(* IEC 61131-3 sources: codesys-motor-control-station/src, 9 files *)

(* ---- types_and_globals.st ---- *)
// ===== E_FaultCode =====

{attribute 'qualified_only'}
{attribute 'strict'}
TYPE E_FaultCode :
(
    NONE     := 0,
    ESTOP    := 1,   // Emergency stop pressed or circuit broken
    OVERLOAD := 2    // Thermal overload relay tripped
) UINT;
END_TYPE

{attribute 'qualified_only'}
{attribute 'strict'}
TYPE E_FaultCode :
(
    NONE     := 0,
    ESTOP    := 1,   // Emergency stop pressed or circuit broken
    OVERLOAD := 2    // Thermal overload relay tripped
) UINT;
END_TYPE

// ===== E_StationState =====

{attribute 'qualified_only'}
{attribute 'strict'}
TYPE E_StationState :
(
    IDLE     := 0,   // Stopped, ready to start
    STARTING := 1,   // Soft-start ramp running
    RUNNING  := 2,   // At speed setpoint
    STOPPING := 3,   // Soft-stop ramp running
    FAULT    := 4    // Fault latched, outputs off
) UINT;
END_TYPE

// ===== ST_Config =====

TYPE ST_Config :
STRUCT
    tRampUp           : TIME := T#5S;    // Soft-start duration (0 Hz to setpoint)
    tRampDown         : TIME := T#5S;    // Soft-stop duration (setpoint to 0 Hz)
    rSpeedMin_Hz      : REAL := 5.0;     // Lowest allowed setpoint
    rSpeedMax_Hz      : REAL := 50.0;    // Highest allowed setpoint
    rSpeedSetpoint_Hz : REAL := 40.0;    // Operator target speed
END_STRUCT
END_TYPE

// ===== GVL_HMI =====

{attribute 'qualified_only'}
VAR_GLOBAL
    xStart        : BOOL;   // Momentary: TRUE while START is pressed
    xStop         : BOOL;   // Momentary: TRUE while STOP is pressed
    xReset        : BOOL;   // Momentary: TRUE while RESET is pressed
    xEStop        : BOOL;   // Latching switch: TRUE = E-stop pressed
    xOverloadTrip : BOOL;   // Latching switch: TRUE = overload tripped
    xSetpointUp   : BOOL;   // Momentary: setpoint +5 Hz
    xSetpointDown : BOOL;   // Momentary: setpoint -5 Hz
END_VAR

// ===== GVL_IO =====

{attribute 'qualified_only'}
VAR_GLOBAL
    // ---------- Inputs ----------
    iEStop_OK       : BOOL;   // NC contact: TRUE = healthy, FALSE = E-stop pressed or wire broken
    iStop_PB        : BOOL;   // NC contact: TRUE = released, FALSE = pressed
    iStart_PB       : BOOL;   // NO contact: TRUE = pressed
    iOverload_OK    : BOOL;   // NC contact: TRUE = healthy, FALSE = overload tripped
    iFaultReset_PB  : BOOL;   // NO contact: TRUE = pressed

    // ---------- Outputs ----------
    qContactor_KM1  : BOOL;   // Main contactor coil
    qDriveRun       : BOOL;   // Run command to the VFD
    qSpeedRef_Hz    : REAL;   // Speed reference sent to the VFD (analog output, in Hz)
    qLamp_Ready     : BOOL;   // White: station ready
    qLamp_Run       : BOOL;   // Green: motor running or ramping
    qLamp_Fault     : BOOL;   // Red: fault latched
END_VAR

// ===== GVL_SIM =====

{attribute 'qualified_only'}
VAR_GLOBAL
    xEnable       : BOOL := TRUE;   // TRUE = simulation writes the GVL_IO inputs

    // Simulated input conditions
    xEStop_OK     : BOOL := TRUE;   // TRUE = E-stop circuit healthy
    xStop_PB      : BOOL := TRUE;   // TRUE = Stop button released
    xStart_PB     : BOOL := FALSE;  // TRUE = Start button pressed
    xOverload_OK  : BOOL := TRUE;   // TRUE = overload circuit healthy
    xFaultReset_PB : BOOL := FALSE; // TRUE = reset button pressed
END_VAR

// ===== GVL_STATION =====

{attribute 'qualified_only'}
VAR_GLOBAL
    stConfig       : ST_Config;                                  // Tunable parameters
    eState         : E_StationState := E_StationState.IDLE;      // Current state machine state
    eFault         : E_FaultCode    := E_FaultCode.NONE;         // Active fault cause
    xFaultLatched  : BOOL;                                       // TRUE until reset
    xSafeToRun     : BOOL;                                       // TRUE only when no fault and all safety inputs healthy
    xRunLatched    : BOOL;                                       // Start/stop seal-in memory
    rSpeedRef_Hz   : REAL;                                       // Ramp output (feeds qSpeedRef_Hz)
    xAtSetpoint    : BOOL;                                       // Ramp has reached the setpoint
    xAtZero        : BOOL;                                       // Ramp has reached 0 Hz
    rRunHours      : REAL;                                       // Run time in hours (for display)
END_VAR

VAR_GLOBAL PERSISTENT RETAIN
    nRunSeconds    : UDINT;                                      // Drive-on time in seconds, survives power cycles
END_VAR

(* ---- FB_RampGenerator.st ---- *)
FUNCTION_BLOCK FB_RampGenerator
VAR_INPUT
    xEnable    : BOOL;              // TRUE = ramp up to target and hold, FALSE = ramp down to 0 Hz
    xForceZero : BOOL;              // TRUE = output jumps to 0 Hz immediately (fault)
    rTarget_Hz : REAL;              // Speed to ramp up to
    tRampUp    : TIME;              // Time to go from 0 Hz to target
    tRampDown  : TIME;              // Time to go from target to 0 Hz
    tCycle     : TIME := T#10MS;    // Task cycle time (must match MainTask)
END_VAR
VAR_OUTPUT
    rOutput_Hz  : REAL;             // Ramped speed reference
    xAtSetpoint : BOOL;             // Enabled and output equals target
    xAtZero     : BOOL;             // Output is 0 Hz
END_VAR
VAR
    rTargetSafe : REAL;             // Target limited to 0 Hz or more
    rGoal       : REAL;             // Where the output is heading right now
    rStepUp     : REAL;             // Hz added per scan while accelerating
    rStepDown   : REAL;             // Hz removed per scan while decelerating
END_VAR
VAR CONSTANT
    rTolerance  : REAL := 0.001;    // Comparison tolerance in Hz
    rMinStep    : REAL := 0.001;    // Smallest allowed step, so a ramp always finishes
END_VAR

// ---------- 1. Goal ----------
rTargetSafe := MAX(rTarget_Hz, 0.0);

IF xEnable THEN
    rGoal := rTargetSafe;
ELSE
    rGoal := 0.0;
END_IF

// ---------- 2. Step sizes per scan ----------
IF tRampUp > T#0S THEN
    rStepUp := MAX(rTargetSafe * TIME_TO_REAL(tCycle) / TIME_TO_REAL(tRampUp), rMinStep);
ELSE
    rStepUp := MAX(rTargetSafe, rMinStep);      // Ramp time 0 = instant
END_IF

IF tRampDown > T#0S THEN
    rStepDown := MAX(rTargetSafe * TIME_TO_REAL(tCycle) / TIME_TO_REAL(tRampDown), rMinStep);
ELSE
    rStepDown := MAX(rTargetSafe, rMinStep);
END_IF

// ---------- 3. Move the output toward the goal ----------
IF xForceZero THEN
    rOutput_Hz := 0.0;
ELSIF rOutput_Hz < rGoal THEN
    rOutput_Hz := MIN(rOutput_Hz + rStepUp, rGoal);
ELSIF rOutput_Hz > rGoal THEN
    rOutput_Hz := MAX(rOutput_Hz - rStepDown, rGoal);
END_IF

// ---------- 4. Status flags ----------
xAtSetpoint := xEnable AND NOT xForceZero AND (ABS(rOutput_Hz - rTargetSafe) <= rTolerance);
xAtZero     := (rOutput_Hz <= rTolerance);

(* ---- PLC_PRG.st ---- *)
PROGRAM PLC_PRG
VAR
    nHeartbeat : UINT;
END_VAR

nHeartbeat := nHeartbeat + 1;   // Proves the task is scanning

PRG_InputSim();                 // 1. Copy simulated and HMI controls to inputs
PRG_Safety();                   // 2. Safety chain
PRG_Station();                  // 3. State machine and outputs
PRG_Ramp();                     // 4. Speed reference ramp
PRG_RunHours();                 // 5. Run-time counter
PRG_HMI();                      // 6. Screen texts and setpoint buttons

(* ---- PRG_HMI.st ---- *)
PROGRAM PRG_HMI
VAR CONSTANT
    rSetpointStep_Hz : REAL := 5.0;     // Change per button click
END_VAR
VAR
    sState   : STRING(30);              // State text for the screen
    sFault   : STRING(30);              // Fault text for the screen
    fbSpUp   : R_TRIG;                  // Edge detect: setpoint up
    fbSpDown : R_TRIG;                  // Edge detect: setpoint down
END_VAR

// ---------- State text ----------
CASE GVL_Station.eState OF
    E_StationState.IDLE:     sState := 'IDLE';
    E_StationState.STARTING: sState := 'STARTING (RAMP UP)';
    E_StationState.RUNNING:  sState := 'RUNNING';
    E_StationState.STOPPING: sState := 'STOPPING (RAMP DOWN)';
    E_StationState.FAULT:    sState := 'FAULT';
END_CASE

// ---------- Fault text ----------
CASE GVL_Station.eFault OF
    E_FaultCode.NONE:     sFault := 'NONE';
    E_FaultCode.ESTOP:    sFault := 'EMERGENCY STOP';
    E_FaultCode.OVERLOAD: sFault := 'MOTOR OVERLOAD';
END_CASE

// ---------- Setpoint buttons (one step per click, kept inside min/max) ----------
fbSpUp  (CLK := GVL_HMI.xSetpointUp);
fbSpDown(CLK := GVL_HMI.xSetpointDown);

IF fbSpUp.Q THEN
    GVL_Station.stConfig.rSpeedSetpoint_Hz := LIMIT(GVL_Station.stConfig.rSpeedMin_Hz,
                                                    GVL_Station.stConfig.rSpeedSetpoint_Hz + rSetpointStep_Hz,
                                                    GVL_Station.stConfig.rSpeedMax_Hz);
END_IF

IF fbSpDown.Q THEN
    GVL_Station.stConfig.rSpeedSetpoint_Hz := LIMIT(GVL_Station.stConfig.rSpeedMin_Hz,
                                                    GVL_Station.stConfig.rSpeedSetpoint_Hz - rSetpointStep_Hz,
                                                    GVL_Station.stConfig.rSpeedMax_Hz);
END_IF

(* ---- PRG_InputSim.st ---- *)
PROGRAM PRG_InputSim
// When enabled, merge the simulator controls and the HMI controls into the project inputs.
// NC contacts (E-stop, Stop, Overload): healthy only if the simulator says healthy AND the HMI is not pressing.
// NO contacts (Start, Reset): active if either source presses.
IF GVL_Sim.xEnable THEN
    GVL_IO.iEStop_OK      := GVL_Sim.xEStop_OK     AND NOT GVL_HMI.xEStop;
    GVL_IO.iStop_PB       := GVL_Sim.xStop_PB      AND NOT GVL_HMI.xStop;
    GVL_IO.iStart_PB      := GVL_Sim.xStart_PB     OR  GVL_HMI.xStart;
    GVL_IO.iOverload_OK   := GVL_Sim.xOverload_OK  AND NOT GVL_HMI.xOverloadTrip;
    GVL_IO.iFaultReset_PB := GVL_Sim.xFaultReset_PB OR GVL_HMI.xReset;
END_IF

(* ---- PRG_Ramp.st ---- *)
PROGRAM PRG_Ramp
VAR CONSTANT
    tTaskCycle : TIME := T#10MS;    // Must equal the MainTask interval
END_VAR
VAR
    fbRamp     : FB_RampGenerator;
    rTarget_Hz : REAL;              // Setpoint limited to the allowed range
END_VAR

// Keep the operator setpoint inside the allowed range
rTarget_Hz := LIMIT(GVL_Station.stConfig.rSpeedMin_Hz,
                    GVL_Station.stConfig.rSpeedSetpoint_Hz,
                    GVL_Station.stConfig.rSpeedMax_Hz);

fbRamp(
    xEnable    := GVL_Station.xRunLatched AND GVL_IO.qDriveRun,   // Ramp starts once the drive has its run command
    xForceZero := NOT GVL_Station.xSafeToRun,                     // Any fault: 0 Hz immediately
    rTarget_Hz := rTarget_Hz,
    tRampUp    := GVL_Station.stConfig.tRampUp,
    tRampDown  := GVL_Station.stConfig.tRampDown,
    tCycle     := tTaskCycle
);

// Publish results
GVL_Station.rSpeedRef_Hz := fbRamp.rOutput_Hz;
GVL_Station.xAtSetpoint  := fbRamp.xAtSetpoint;
GVL_Station.xAtZero      := fbRamp.xAtZero;

// Analog output to the VFD
GVL_IO.qSpeedRef_Hz := GVL_Station.rSpeedRef_Hz;

(* ---- PRG_RunHours.st ---- *)
PROGRAM PRG_RunHours
VAR CONSTANT
    nTaskCycle_ms : UDINT := 10;    // Must equal the MainTask interval
END_VAR
VAR
    nMilliseconds : UDINT;          // Partial second, carried over between runs
END_VAR

// Count time while the VFD run command is active (includes the stop ramp)
IF GVL_IO.qDriveRun THEN
    nMilliseconds := nMilliseconds + nTaskCycle_ms;

    IF nMilliseconds >= 1000 THEN
        nMilliseconds := nMilliseconds - 1000;
        GVL_Station.nRunSeconds := GVL_Station.nRunSeconds + 1;
    END_IF
END_IF

GVL_Station.rRunHours := UDINT_TO_REAL(GVL_Station.nRunSeconds) / 3600.0;

(* ---- PRG_Safety.st ---- *)
PROGRAM PRG_Safety
VAR
    fbResetTrig     : R_TRIG;   // Detects the rising edge of the reset button
    xEStopActive    : BOOL;     // TRUE while E-stop circuit is open
    xOverloadActive : BOOL;     // TRUE while overload relay is tripped
    xResetAllowed   : BOOL;     // TRUE when a latched fault may be cleared
END_VAR

// ---------- 1. Raw conditions (NC inputs: FALSE means a problem) ----------
xEStopActive    := NOT GVL_IO.iEStop_OK;
xOverloadActive := NOT GVL_IO.iOverload_OK;

// ---------- 2. Fault latch (E-stop has priority over overload) ----------
IF xEStopActive THEN
    GVL_Station.xFaultLatched := TRUE;
    GVL_Station.eFault        := E_FaultCode.ESTOP;
ELSIF xOverloadActive AND NOT GVL_Station.xFaultLatched THEN
    GVL_Station.xFaultLatched := TRUE;
    GVL_Station.eFault        := E_FaultCode.OVERLOAD;
END_IF

// ---------- 3. Fault reset (edge-triggered, only when the cause is gone) ----------
fbResetTrig(CLK := GVL_IO.iFaultReset_PB);
xResetAllowed := GVL_Station.xFaultLatched AND NOT xEStopActive AND NOT xOverloadActive;

IF fbResetTrig.Q AND xResetAllowed THEN
    GVL_Station.xFaultLatched := FALSE;
    GVL_Station.eFault        := E_FaultCode.NONE;
END_IF

// ---------- 4. Permissive for the rest of the program ----------
GVL_Station.xSafeToRun := NOT GVL_Station.xFaultLatched
                          AND NOT xEStopActive
                          AND NOT xOverloadActive;

(* ---- PRG_Station.st ---- *)
PROGRAM PRG_Station
VAR CONSTANT
    tContactorDelay : TIME := T#500MS;   // Wait after KM1 closes before the drive gets its run command
    tBlinkHalf      : TIME := T#500MS;   // Half period of the lamp blinker
END_VAR
VAR
    fbStartTrig   : R_TRIG;   // Rising edge of the Start button
    fbDriveDelay  : TON;      // Contactor pull-in delay
    fbBlink       : TON;      // Blink generator
    xBlink        : BOOL;     // 1 Hz blink signal
    xMotorPowered : BOOL;     // TRUE when the contactor should be closed
END_VAR

// ---------- 1. Start/stop seal-in ----------
// Start: NO button, accepted only in IDLE on a rising edge.
// Stop: NC button (TRUE = released). Stop and safety always win.
fbStartTrig(CLK := GVL_IO.iStart_PB);

GVL_Station.xRunLatched := (   (fbStartTrig.Q AND (GVL_Station.eState = E_StationState.IDLE))
                            OR GVL_Station.xRunLatched )
                           AND GVL_IO.iStop_PB
                           AND GVL_Station.xSafeToRun;

// ---------- 2. State machine ----------
IF NOT GVL_Station.xSafeToRun THEN
    GVL_Station.eState := E_StationState.FAULT;
ELSE
    CASE GVL_Station.eState OF

        E_StationState.FAULT:
            // Safety is healthy again (fault was reset)
            GVL_Station.eState := E_StationState.IDLE;

        E_StationState.IDLE:
            IF GVL_Station.xRunLatched THEN
                GVL_Station.eState := E_StationState.STARTING;
            END_IF

        E_StationState.STARTING:
            IF NOT GVL_Station.xRunLatched THEN
                GVL_Station.eState := E_StationState.STOPPING;
            ELSIF GVL_Station.xAtSetpoint THEN
                GVL_Station.eState := E_StationState.RUNNING;
            END_IF

        E_StationState.RUNNING:
            IF NOT GVL_Station.xRunLatched THEN
                GVL_Station.eState := E_StationState.STOPPING;
            END_IF

        E_StationState.STOPPING:
            IF GVL_Station.xAtZero THEN
                GVL_Station.eState := E_StationState.IDLE;
            END_IF

    END_CASE
END_IF

// ---------- 3. Contactor and drive run command ----------
xMotorPowered := (GVL_Station.eState = E_StationState.STARTING)
              OR (GVL_Station.eState = E_StationState.RUNNING)
              OR (GVL_Station.eState = E_StationState.STOPPING);

GVL_IO.qContactor_KM1 := xMotorPowered;

fbDriveDelay(IN := xMotorPowered, PT := tContactorDelay);
GVL_IO.qDriveRun := fbDriveDelay.Q;

// ---------- 4. Lamps ----------
// Blink generator: the TON restarts itself, giving one pulse every tBlinkHalf
fbBlink(IN := NOT fbBlink.Q, PT := tBlinkHalf);
IF fbBlink.Q THEN
    xBlink := NOT xBlink;
END_IF

GVL_IO.qLamp_Ready := (GVL_Station.eState = E_StationState.IDLE);

GVL_IO.qLamp_Run   := (GVL_Station.eState = E_StationState.RUNNING)
                      OR ( xBlink AND (    (GVL_Station.eState = E_StationState.STARTING)
                                        OR (GVL_Station.eState = E_StationState.STOPPING) ) );

GVL_IO.qLamp_Fault := GVL_Station.xFaultLatched;
